(* IEC 61131-3 sources: llm-plc-st-eval/data/calibracion/claude-sonnet-4-6/A6/few_shot, 3 files *)

(* ---- ejec_1.st ---- *)
```st
FUNCTION_BLOCK FB_Modos
VAR_INPUT
    selector       : INT;                  (* Selector de modo: 0=Auto, 1=Manual, 2=Mantenimiento *)
    estadoSeguro   : BOOL;                 (* Permiso para cambiar modo y mantener forzados *)
    cmdAuto        : ARRAY[0..7] OF BOOL;  (* Comandos en modo automatico *)
    cmdManual      : ARRAY[0..7] OF BOOL;  (* Comandos en modo manual *)
    idxForzado     : INT;                  (* Indice del actuador a forzar (0-7) *)
    valorForzado   : BOOL;                 (* Valor a aplicar al actuador forzado *)
    confirmarForzado : BOOL;               (* Flanco ascendente aplica el forzado *)
END_VAR
VAR_OUTPUT
    modoActivo : INT;                      (* Modo vigente: 0=Auto, 1=Manual, 2=Mantenimiento *)
    actuador   : ARRAY[0..7] OF BOOL;      (* Estado de los ocho actuadores *)
END_VAR
VAR
    prevConfirmar  : BOOL;                 (* Valor anterior de confirmarForzado para deteccion de flanco *)
    estadoForzado  : ARRAY[0..7] OF BOOL;  (* Valores forzados en modo mantenimiento *)
    prevEstadoSeguro : BOOL;               (* Valor anterior de estadoSeguro *)
    i              : INT;                  (* Indice de iteracion *)
    primerCiclo    : BOOL := TRUE;         (* Bandera de primer ciclo para inicializacion *)
END_VAR

(* --- Inicializacion en el primer ciclo: modo manual por defecto --- *)
IF primerCiclo THEN
    modoActivo   := 1;
    primerCiclo  := FALSE;
END_IF;

(* --- Gestion del cambio de modo --- *)
(* Solo se acepta un selector valido (0-2) cuando estadoSeguro esta activo *)
IF estadoSeguro THEN
    IF selector >= 0 AND selector <= 2 THEN
        IF selector <> modoActivo THEN
            (* Al salir de mantenimiento se anulan todos los forzados *)
            IF modoActivo = 2 THEN
                FOR i := 0 TO 7 DO
                    estadoForzado[i] := FALSE;
                END_FOR;
            END_IF;
            modoActivo := selector;
        END_IF;
    END_IF;
    (* Valores fuera de rango se ignoran: modoActivo no cambia *)
END_IF;

(* --- Mantenimiento: si estadoSeguro se desactiva, apagar todos los actuadores forzados --- *)
IF modoActivo = 2 THEN
    IF NOT estadoSeguro AND prevEstadoSeguro THEN
        (* Flanco descendente de estadoSeguro durante mantenimiento *)
        FOR i := 0 TO 7 DO
            estadoForzado[i] := FALSE;
        END_FOR;
    END_IF;

    (* Aplicar forzado en flanco ascendente de confirmarForzado, solo si estadoSeguro activo *)
    IF confirmarForzado AND NOT prevConfirmar THEN
        IF estadoSeguro THEN
            IF idxForzado >= 0 AND idxForzado <= 7 THEN
                estadoForzado[idxForzado] := valorForzado;
            END_IF;
            (* idxForzado fuera de rango se ignora *)
        END_IF;
    END_IF;
END_IF;

(* --- Actualizacion de salidas segun modo vigente --- *)
CASE modoActivo OF
    0: (* Automatico: cada actuador sigue a cmdAuto *)
        FOR i := 0 TO 7 DO
            actuador[i] := cmdAuto[i];
        END_FOR;

    1: (* Manual: cada actuador sigue a cmdManual *)
        FOR i := 0 TO 7 DO
            actuador[i] := cmdManual[i];
        END_FOR;

    2: (* Mantenimiento: actuadores reflejan los forzados (apagados si no se han forzado) *)
        FOR i := 0 TO 7 DO
            actuador[i] := estadoForzado[i];
        END_FOR;
END_CASE;

(* --- Guardar valores previos para proxima ejecucion --- *)
prevConfirmar    := confirmarForzado;
prevEstadoSeguro := estadoSeguro;

END_FUNCTION_BLOCK
```

(* ---- ejec_2.st ---- *)
```structured-text
FUNCTION_BLOCK FB_Modos
VAR_INPUT
    selector       : INT;                  (* Selector de modo: 0=Auto, 1=Manual, 2=Mantenimiento *)
    estadoSeguro   : BOOL;                 (* Permiso para cambio de modo y forzados *)
    cmdAuto        : ARRAY[0..7] OF BOOL;  (* Comandos en modo automatico *)
    cmdManual      : ARRAY[0..7] OF BOOL;  (* Comandos en modo manual *)
    idxForzado     : INT;                  (* Indice del actuador a forzar en mantenimiento *)
    valorForzado   : BOOL;                 (* Valor a aplicar al actuador forzado *)
    confirmarForzado : BOOL;               (* Flanco ascendente aplica el forzado *)
END_VAR
VAR_OUTPUT
    modoActivo : INT;                      (* Modo vigente: 0=Auto, 1=Manual, 2=Mantenimiento *)
    actuador   : ARRAY[0..7] OF BOOL;      (* Estado de los ocho actuadores *)
END_VAR
VAR
    prevConfirmar  : BOOL;                 (* Valor anterior de confirmarForzado para deteccion de flanco *)
    prevSeguro     : BOOL;                 (* Valor anterior de estadoSeguro *)
    forzados       : ARRAY[0..7] OF BOOL;  (* Valores forzados en modo mantenimiento *)
    i              : INT;                  (* Indice de iteracion *)
    flancoCon      : BOOL;                 (* Flanco ascendente de confirmarForzado *)
    flancoSeguro   : BOOL;                 (* Flanco ascendente de estadoSeguro *)
    primeraEjecucion : BOOL;              (* Bandera de inicializacion *)
END_VAR

(* ── Inicializacion en la primera ejecucion ── *)
IF NOT primeraEjecucion THEN
    modoActivo       := 1;   (* Modo inicial: manual *)
    primeraEjecucion := TRUE;
    prevConfirmar    := FALSE;
    prevSeguro       := estadoSeguro;
END_IF;

(* ── Deteccion de flancos ── *)
flancoCon    := confirmarForzado AND NOT prevConfirmar;
flancoSeguro := estadoSeguro AND NOT prevSeguro;

(* ── Gestion del cambio de modo ── *)
(* Se acepta un nuevo modo si estadoSeguro esta activo y el selector es valido (0..2) *)
IF estadoSeguro AND (selector >= 0) AND (selector <= 2) AND (selector <> modoActivo) THEN
    (* Al salir de mantenimiento se anulan todos los forzados *)
    IF modoActivo = 2 THEN
        FOR i := 0 TO 7 DO
            forzados[i] := FALSE;
        END_FOR;
    END_IF;
    modoActivo := selector;
END_IF;

(* ── Logica de modo mantenimiento ── *)
IF modoActivo = 2 THEN
    (* Si estadoSeguro se desactiva durante mantenimiento, apagar y anular forzados *)
    IF NOT estadoSeguro THEN
        FOR i := 0 TO 7 DO
            forzados[i] := FALSE;
            actuador[i] := FALSE;
        END_FOR;
    ELSE
        (* Aplicar forzado en flanco ascendente de confirmarForzado con indice valido *)
        IF flancoCon AND (idxForzado >= 0) AND (idxForzado <= 7) THEN
            forzados[idxForzado] := valorForzado;
        END_IF;
        (* Los actuadores reflejan los valores forzados *)
        FOR i := 0 TO 7 DO
            actuador[i] := forzados[i];
        END_FOR;
    END_IF;

(* ── Logica de modo automatico ── *)
ELSIF modoActivo = 0 THEN
    FOR i := 0 TO 7 DO
        actuador[i] := cmdAuto[i];
    END_FOR;

(* ── Logica de modo manual ── *)
ELSE (* modoActivo = 1 *)
    FOR i := 0 TO 7 DO
        actuador[i] := cmdManual[i];
    END_FOR;
END_IF;

(* ── Actualizacion de valores previos ── *)
prevConfirmar := confirmarForzado;
prevSeguro    := estadoSeguro;

END_FUNCTION_BLOCK
```

(* ---- ejec_3.st ---- *)
```st
FUNCTION_BLOCK FB_Modos
VAR_INPUT
    selector       : INT;                  (* Modo deseado: 0=Auto, 1=Manual, 2=Mant. *)
    estadoSeguro   : BOOL;                 (* Permiso para cambiar modo y forzar *)
    cmdAuto        : ARRAY[0..7] OF BOOL;  (* Comandos en modo automatico *)
    cmdManual      : ARRAY[0..7] OF BOOL;  (* Comandos en modo manual *)
    idxForzado     : INT;                  (* Indice del actuador a forzar *)
    valorForzado   : BOOL;                 (* Valor a aplicar al actuador forzado *)
    confirmarForzado : BOOL;               (* Flanco ascendente aplica el forzado *)
END_VAR
VAR_OUTPUT
    modoActivo : INT;                      (* Modo vigente: 0=Auto, 1=Manual, 2=Mant. *)
    actuador   : ARRAY[0..7] OF BOOL;     (* Estado de los ocho actuadores *)
END_VAR
VAR
    i                  : INT;             (* Indice de iteracion *)
    prevConfirmar      : BOOL;            (* Valor anterior de confirmarForzado *)
    prevEstadoSeguro   : BOOL;            (* Valor anterior de estadoSeguro *)
    estadosForzados    : ARRAY[0..7] OF BOOL; (* Valores forzados en mantenimiento *)
    primerCiclo        : BOOL := TRUE;    (* Marca de primer ciclo para inicializacion *)
END_VAR

(* ── Inicializacion en el primer ciclo: modo manual ── *)
IF primerCiclo THEN
    modoActivo  := 1;
    primerCiclo := FALSE;
END_IF;

(* ── Gestion de cambio de modo ── *)
(* Solo se acepta un selector valido (0..2) cuando estadoSeguro esta activo *)
IF estadoSeguro AND (selector >= 0) AND (selector <= 2) THEN
    IF selector <> modoActivo THEN
        (* Al salir de mantenimiento, anular todos los forzados *)
        IF modoActivo = 2 THEN
            FOR i := 0 TO 7 DO
                estadosForzados[i] := FALSE;
            END_FOR;
        END_IF;
        modoActivo := selector;
    END_IF;
END_IF;

(* ── Logica especifica de mantenimiento ── *)
IF modoActivo = 2 THEN

    (* Si estadoSeguro se desactiva durante mantenimiento: apagar y anular forzados *)
    IF prevEstadoSeguro AND NOT estadoSeguro THEN
        FOR i := 0 TO 7 DO
            estadosForzados[i] := FALSE;
        END_FOR;
    END_IF;

    (* Detectar flanco ascendente de confirmarForzado *)
    IF confirmarForzado AND NOT prevConfirmar THEN
        (* Solo si estadoSeguro activo e indice valido *)
        IF estadoSeguro AND (idxForzado >= 0) AND (idxForzado <= 7) THEN
            estadosForzados[idxForzado] := valorForzado;
        END_IF;
    END_IF;

END_IF;

(* ── Actualizacion de salidas de actuadores ── *)
FOR i := 0 TO 7 DO
    CASE modoActivo OF
        0: (* Automatico *)
            actuador[i] := cmdAuto[i];
        1: (* Manual *)
            actuador[i] := cmdManual[i];
        2: (* Mantenimiento *)
            IF estadoSeguro THEN
                actuador[i] := estadosForzados[i];
            ELSE
                actuador[i] := FALSE; (* Sin estado seguro, todo apagado *)
            END_IF;
    ELSE
        actuador[i] := FALSE; (* Modo desconocido: seguridad *)
    END_CASE;
END_FOR;

(* ── Guardar valores previos para proximos ciclos ── *)
prevConfirmar    := confirmarForzado;
prevEstadoSeguro := estadoSeguro;

END_FUNCTION_BLOCK
```
